(* IEC 61131-3 sources: SRCI_CLIENT_PLC/RobotLibrary/Library/POUs/Additional/MC_OpenBrake/Structures, 4 files *)

(* ---- OpenBrakeOutCmd.st ---- *)
{attribute 'pack_mode' := '1'}
// -------------------------------------------------------------------------
//  SRCI Robot Library
// -------------------------------------------------------------------------
//
//  Object:      BrakeTestOutCmd
//  Author:      Thorsten Brach
//  Date:        2024-06-01
//
//  Description:
//
//
//  Copyright:
//    (C) 2024 Thorsten Brach. All rights reserved
//             Licensed under the MIT License.
//
//  Disclaimer:
//    This project is provided without any guarantee and can be used for
//    private and commercial purposes. Any use is at the user’s
//    own risk and responsibility.
//
// -------------------------------------------------------------------------
TYPE OpenBrakeOutCmd :
STRUCT
  /// TRUE when "OpenBrake" is active.
  Enabled                   : BOOL;
  /// Indicates the brake release status of the main robot axes.
  /// • TRUE: The brake of the axis is opened.
  /// • FALSE: The brake of the axis is closed.
  /// See Table 6-698 for bit assignment
  RobotAxesBrakeReleased    : RobotAxesFlags;
  /// Indicates the brake release status of the external robot axes.
  /// • TRUE: The brake of the axis is opened.
  /// • FALSE: The brake of the axis is closed/not supported
  /// See Table 6-698 for bit assignment
  ExternalAxesBrakeReleased : ExternalAxesFlags;
END_STRUCT
END_TYPE

(* ---- OpenBrakeParCmd.st ---- *)
{attribute 'pack_mode' := '1'}
// -------------------------------------------------------------------------
//  SRCI Robot Library
// -------------------------------------------------------------------------
//
//  Object:      OpenBrakeParCmd
//  Author:      Thorsten Brach
//  Date:        2024-06-01
//
//  Description:
//
//
//  Copyright:
//    (C) 2024 Thorsten Brach. All rights reserved
//             Licensed under the MIT License.
//
//  Disclaimer:
//    This project is provided without any guarantee and can be used for
//    private and commercial purposes. Any use is at the user’s
//    own risk and responsibility.
//
// -------------------------------------------------------------------------
TYPE OpenBrakeParCmd :
STRUCT
  /// Defines which brake of the robot axes must be released.
  /// • TRUE: Open the brake of the axis.
  /// • FALSE (default): Close the brake of the axis.
  RobotAxesBrakeRelease    : RobotAxesFlags;
  /// Defines which brake of the external robot axis must be released.
  /// • TRUE: Open the brake of the axis.
  /// • FALSE (default): Close the brake of the axis.
  /// See Table 6-698 for bit assignment.
  ExternalAxesBrakeRelease : ExternalAxesFlags;
END_STRUCT
END_TYPE

(* ---- OpenBrakeRecvData.st ---- *)
{attribute 'pack_mode' := '1'}
// -------------------------------------------------------------------------
//  SRCI Robot Library
// -------------------------------------------------------------------------
//
//  Object:      BrakeTestRecvData
//  Author:      Thorsten Brach
//  Date:        2024-06-01
//
//  Description:
//
//
//  Copyright:
//    (C) 2024 Thorsten Brach. All rights reserved
//             Licensed under the MIT License.
//
//  Disclaimer:
//    This project is provided without any guarantee and can be used for
//    private and commercial purposes. Any use is at the user’s
//    own risk and responsibility.
//
// -------------------------------------------------------------------------
TYPE OpenBrakeRecvData EXTENDS RspHeader :
STRUCT
  /// TRUE when "OpenBrake" is active.
  Enabled                   : BYTE;
  /// Indicates the brake release status of the main robot axes.
  /// • TRUE: The brake of the axis is opened.
  /// • FALSE: The brake of the axis is closed.
  /// See Table 6-698 for bit assignment
  RobotAxesBrakeReleased    : BYTE;
  /// Indicates the brake release status of the external robot axes.
  /// • TRUE: The brake of the axis is opened.
  /// • FALSE: The brake of the axis is closed/not supported
  /// See Table 6-698 for bit assignment
  ExternalAxesBrakeReleased : BYTE;
END_STRUCT
END_TYPE

(* ---- OpenBrakeSendData.st ---- *)
{attribute 'pack_mode' := '1'}
// -------------------------------------------------------------------------
//  SRCI Robot Library
// -------------------------------------------------------------------------
//
//  Object:      BrakeTestSendData
//  Author:      Thorsten Brach
//  Date:        2024-06-01
//
//  Description:
//
//
//  Copyright:
//    (C) 2024 Thorsten Brach. All rights reserved
//             Licensed under the MIT License.
//
//  Disclaimer:
//    This project is provided without any guarantee and can be used for
//    private and commercial purposes. Any use is at the user’s
//    own risk and responsibility.
//
// -------------------------------------------------------------------------
TYPE OpenBrakeSendData EXTENDS CmdHeader:
STRUCT
  /// Defines which brake of the robot axes must be released.
  /// • TRUE: Open the brake of the axis.
  /// • FALSE (default): Close the brake of the axis.
  RobotAxesBrakeRelease    : BYTE;
  /// Defines which brake of the external robot axis must be released.
  /// • TRUE: Open the brake of the axis.
  /// • FALSE (default): Close the brake of the axis.
  /// See Table 6-698 for bit assignment.
  ExternalAxesBrakeRelease : BYTE;
END_STRUCT
END_TYPE
